ABB RobotStudio station: 项目1.rsstn

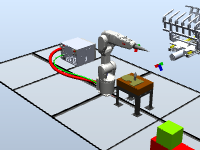
Station Station (saved by RobotStudio 6.8.8148.134)
Controller System1
  mechanical unit ROB_1: ?, 6 joints, base frame (0, 0, 0) mm
Layout (positions relative to the parent item):
  - IRB1200_5_90_STD_02 [mechanism, from Robots\IRB1200_5_90_STD_02.rslib] at (0, 0, 0) mm; joint values [0, 0, 0, 0, 0, 0] (rad or m)
  - IRC5_Compact [part, from Equipment\IRC5_Compact__02.rslib] at (-1416.87, 226.47, 0) mm
  - table_and_fixture_140 [part, from Training Objects\propeller_table.rslib] at (317.24, -175, 0) mm
  - 圆锥 [part]
  - PhysicsCable_1 [physicscable]
  - PhysicsCable_3 [physicscable]
  - 部件_2 [part] at (0, 0, 718.85) mm, rotated rx 180 ry 0 rz 0 deg
  - 轨道 [mechanism] at (1267.8, -633.39, 2.84) mm; joint values [0.0756] (rad or m)
      links: L1, L2
  - 夹具 [mechanism] at (0, 0, 694.72) mm; joint values [0.6934] (rad or m)
      links: L1, L2, L3
  - Curve_thing [part, from Training Objects\Curve_Thing.rslib] at (342.24, -150, 308) mm
  - 部件_3 [part] at (533, 0, 889.1) mm, rotated rx 0 ry 90 rz 0 deg
Attachment: 部件_3 is attached to IRB1200_5_90_STD_02 / Link6
Targets, tools, work objects and paths stored in the station, written as RAPID:
! task (no controller)
MODULE CalibData
  PERS tooldata tWeldGun:=[TRUE,[[125.800591275,0,391.268161315],[0.898794046,0,0.438371147,0]],[3,[0,0,100],[0,1,0,0],0,0,0]];
ENDMODULE

